(* IEC 61131-3 sources: kns-port-domestic/tools/plcopen/tests/fixtures/constructs/src/POUs/Devices/FB_Motor, 8 files *)

(* ---- FB_Motor.decl.st ---- *)
// Назначение: двигатель — наследник базы: пуск, сброс через SUPER^, счёт пусков
// Автор:      <ИМЯ ФАМИЛИЯ>
// Версия:     0.1.0
// Документ:   docs/plcopen.md
FUNCTION_BLOCK FB_Motor EXTENDS FB_DeviceBase
VAR_INPUT
    stCmd : ST_MotorCmd;
END_VAR
VAR_OUTPUT
    xRun : BOOL;
END_VAR
VAR
    uiStarts : UINT;
    fbCounter : FB_Counter;
END_VAR

(* ---- Describe.method.decl.st ---- *)
// Описание для журнала
METHOD PRIVATE FINAL Describe : WSTRING(40)
VAR
    wsText : WSTRING(40) := "Двигатель";
END_VAR

(* ---- FB_init.method.decl.st ---- *)
// Инициализация экземпляра
METHOD FB_init : BOOL
VAR_INPUT
    bInitRetains : BOOL;    // TRUE — инициализировать RETAIN
    bInCopyCode : BOOL;     // TRUE — экземпляр копируется при онлайн-изменении
END_VAR

(* ---- FB_Motor.impl.st ---- *)
SUPER^();
IF stCmd.xStart AND NOT xFault THEN
    Start();
ELSIF stCmd.xStop THEN
    xRun := FALSE;
END_IF

(* ---- Reset.method.decl.st ---- *)
METHOD PUBLIC Reset : BOOL
VAR_INPUT
    xForce : BOOL;
END_VAR

(* ---- Start.method.decl.st ---- *)
METHOD PUBLIC Start : BOOL
VAR_INST
    uiCalls : UINT;     // число вызовов метода (сохраняется между вызовами)
END_VAR

(* ---- Start.method.impl.st ---- *)
uiCalls := uiCalls + 1;
IF THIS^.Mode = E_Mode.Auto OR Mode = E_Mode.Manual THEN
    xRun := TRUE;
    uiStarts := uiStarts + 1;
END_IF
Start := xRun;

(* ---- Starts.get.decl.st ---- *)
VAR
    uiCopy : UINT;
END_VAR
